(* IEC 61131-3 sources: kns-port-domestic/tools/plcopen/tests/fixtures/constructs/src/DUTs, 7 files *)

(* ---- E_Color.dut.st ---- *)
// Перечисление без значений и без базового типа
TYPE E_Color :
(
    Red,
    Green,
    Blue
);
END_TYPE

(* ---- E_Mode.dut.st ---- *)
// Режим устройства: перечисление с явными значениями и базовым типом
{attribute 'qualified_only'}
{attribute 'strict'}
TYPE E_Mode :
(
    OutOfService := 0,  // выведено из работы
    Auto := 1,          // автоматический
    Manual := 2,        // ручной
    Local := 3          // местный
) INT;
END_TYPE

(* ---- ST_Base.dut.st ---- *)
// Базовая структура: начальные значения, массив, строка, комментарии
TYPE ST_Base :
STRUCT
    xEnable : BOOL := TRUE;               // разрешение
    iCount : INT;                         (* счётчик *)
    rValue_bar : REAL := 1.5;
    sName : STRING(32) := 'base';
    wsLabel : WSTRING(16) := "Насос";
    aiData : ARRAY[0..3] OF INT := [1, 2, 3, 4];
    eMode : E_Mode := E_Mode.Auto;
END_STRUCT
END_TYPE

(* ---- ST_Derived.dut.st ---- *)
// Структура-наследник базовой
TYPE ST_Derived EXTENDS ST_Base :
STRUCT
    tDelay : TIME := T#5S;
    ltStamp : LTIME;
    pData : POINTER TO INT;
END_STRUCT
END_TYPE

(* ---- T_Name.dut.st ---- *)
// Псевдоним строкового типа
TYPE T_Name : STRING(20);
END_TYPE

(* ---- T_Percent.dut.st ---- *)
// Псевдоним с поддиапазоном
TYPE T_Percent : INT(0..100);
END_TYPE

(* ---- U_Raw.dut.st ---- *)
// Объединение: одно слово как целое и как биты
TYPE U_Raw :
UNION
    wWord : WORD;
    aBytes : ARRAY[0..1] OF BYTE;
END_UNION
END_TYPE
